{attribute 'qualified_only'}
VAR_GLOBAL CONSTANT
	cMaxArguments		: USINT := 10;				// placeholders {0}..{9}
	cLanguageCount		: USINT := 11;				// number of values in E_Language - raise when adding a language
	HR_NO_CONTEXT		: HRESULT := -2147467261;	// 16#80004003 (E_POINTER): no I_EventContext was injected
	HR_NOT_IMPLEMENTED	: HRESULT := -2147467263;	// 16#80004001 (E_NOTIMPL)
END_VAR

(* stored: Version 1.1.0.1
   GVL GVL_EventFramework: Id {b0f33a38-8cac-420c-968b-7d54139b9f8d} *)
